// TIA Portal V20 export
Screen "Pop-up_PLP"  472x499
  ScreenItem "Background" at 0,0 size 472x499  Type=HmiRectangle
  ScreenItem "Rectangle TG Status" at 0,1 size 372x43  Type=HmiRectangle
  ScreenItem "Rectangle TG1" at 0,31 size 372x55  Type=HmiRectangle
  ScreenItem "Text Field TG1 In Pounce Pos" at 186,36 size 90x21  Type=HmiTextBox
  ScreenItem "Text Field TG1 In Work Pos" at 275,36 size 90x21  Type=HmiTextBox
  ScreenItem "Text field TG1 Status" at 8,62 size 47x21  Type=HmiTextBox
  ScreenItem "Text Field TG1 Fault" at 8,36 size 90x21  Type=HmiTextBox
  ScreenItem "Text Field TG1 In Home Pos" at 97,36 size 90x21  Type=HmiTextBox
  ScreenItem "Rectangle TG2" at 0,86 size 372x55  Type=HmiRectangle
  ScreenItem "Text Field TG2 In Pounce Pos" at 186,91 size 90x21  Type=HmiTextBox
  ScreenItem "Text Field TG2 In Work Pos" at 275,91 size 90x21  Type=HmiTextBox
  ScreenItem "Text field TG2 Status" at 8,116 size 47x21  Type=HmiTextBox
  ScreenItem "Text Field TG2 Fault" at 8,91 size 90x21  Type=HmiTextBox
  ScreenItem "Text Field TG2 In Home Pos" at 97,91 size 90x21  Type=HmiTextBox
  ScreenItem "Rectangle TG3" at 0,141 size 372x55  Type=HmiRectangle
  ScreenItem "Text Field TG3 In Pounce Pos" at 186,146 size 90x21  Type=HmiTextBox
  ScreenItem "Text Field TG3 In Work Pos" at 275,146 size 90x21  Type=HmiTextBox
  ScreenItem "Text field TG3 Status" at 8,171 size 47x21  Type=HmiTextBox
  ScreenItem "Text Field TG3 Fault" at 8,146 size 90x21  Type=HmiTextBox
  ScreenItem "Text Field TG3 In Home Pos" at 97,146 size 90x21  Type=HmiTextBox
  ScreenItem "Rectangle TG4" at 0,196 size 372x55  Type=HmiRectangle
  ScreenItem "Text Field TG4 In Pounce Pos" at 186,201 size 90x21  Type=HmiTextBox
  ScreenItem "Text Field TG4 In Work Pos" at 275,201 size 90x21  Type=HmiTextBox
  ScreenItem "Text field TG4 Status" at 8,227 size 47x21  Type=HmiTextBox
  ScreenItem "Text Field TG4 Fault" at 8,201 size 90x21  Type=HmiTextBox
  ScreenItem "Text Field TG4 In Home Pos" at 97,201 size 90x21  Type=HmiTextBox
  ScreenItem "Rectangle TG5" at 0,251 size 372x55  Type=HmiRectangle
  ScreenItem "Text Field TG5 In Pounce Pos" at 186,256 size 90x21  Type=HmiTextBox
  ScreenItem "Text Field TG5 In Work Pos" at 275,256 size 90x21  Type=HmiTextBox
  ScreenItem "Text field TG5 Status" at 8,281 size 47x21  Type=HmiTextBox
  ScreenItem "Text Field TG5 Fault" at 8,256 size 90x21  Type=HmiTextBox
  ScreenItem "Text Field TG5 In Home Pos" at 97,256 size 90x21  Type=HmiTextBox
  ScreenItem "Rectangle TG6" at 0,306 size 372x55  Type=HmiRectangle
  ScreenItem "Text Field TG6 In Pounce Pos" at 186,311 size 90x21  Type=HmiTextBox
  ScreenItem "Text Field TG6 In Work Pos" at 275,311 size 90x21  Type=HmiTextBox
  ScreenItem "Text field TG6 Status" at 8,336 size 47x21  Type=HmiTextBox
  ScreenItem "Text Field TG6 Fault" at 8,311 size 90x21  Type=HmiTextBox
  ScreenItem "Text Field TG6 In Home Pos" at 97,311 size 90x21  Type=HmiTextBox
  ScreenItem "Rectangle TG7" at 0,361 size 372x55  Type=HmiRectangle
  ScreenItem "Text Field TG7 In Pounce Pos" at 186,366 size 90x21  Type=HmiTextBox
  ScreenItem "Text Field TG7 In Work Pos" at 275,366 size 90x21  Type=HmiTextBox
  ScreenItem "Text field TG7 Status" at 8,392 size 47x21  Type=HmiTextBox
  ScreenItem "Text Field TG7 Fault" at 8,366 size 90x21  Type=HmiTextBox
  ScreenItem "Text Field TG7 In Home Pos" at 97,366 size 90x21  Type=HmiTextBox
  ScreenItem "Rectangle TG8" at 0,416 size 372x55  Type=HmiRectangle
  ScreenItem "Text Field TG8 In Pounce Pos" at 186,421 size 90x21  Type=HmiTextBox
  ScreenItem "Text Field TG8 In Work Pos" at 275,421 size 90x21  Type=HmiTextBox
  ScreenItem "Text field TG8 Status" at 8,446 size 47x21  Type=HmiTextBox
  ScreenItem "Text Field TG8 Fault" at 8,421 size 90x21  Type=HmiTextBox
  ScreenItem "Text Field TG8 In Home Pos" at 97,421 size 90x21  Type=HmiTextBox
  ScreenItem "Text field TG Status" at 0,0 size 373x31  Type=HmiTextBox
  ScreenItem "Move_Legend" at 382,0 size 90x60  Type=HmiButton
